SUBAPPLICATION logiBUS_PI_Speed_Publish_OPC (* logiBUS_PI_IDA (Puls-Eingang) als Frequenz (Hz, nur lokal fuer Dashboard/Diagnose) UND als bereits auf die physikalische Einheit umgerechneter Endwert (SCALE+RASTER, M2M-Publish fuer andere Stationen) ausgeben - OHNE jegliche VT-Interaktion. Erweiterung von logiBUS_PI_Raw_Publish_OPC um die Hz->Einheit-Umrechnung (bisher zentral auf STG1 via AR_HZ_TO_Q_Publish_OPC) - jetzt co-located mit dem Sensor: nur der fertige physikalische Endwert verlaesst die Station M2M, der rohe Hz-Wert bleibt lokal. *)
  (* Standard: 61499-2; Description: Copyright (c) 2026 Meisterschulen am Ostbahnhof This program and the accompanying materials are made available under the terms of the Eclipse Public License 2.0 which is available at https://www.eclipse.org/legal/epl-2.0/ SPDX-License-Identifier: EPL-2.0 *)
  (* Version 1.3, 2026-10-03, Franz Höpfinger, Meisterschulen am Ostbahnhof, Franz: 'K auch auf Adapter umstellen' - FT_DERIV_10_AR.K ist jetzt selbst ein AUI-Adapter-Socket (FT_DERIV_10_AR v1.2), die bisherige Entpack-Umgehung ToUINT (AUI_UI_TO_UINT) entfaellt dadurch ersatzlos: ToAUI.AUI_OUT verdrahtet jetzt direkt auf FT_DERIV_10_AR.K (beides AUI-Adapter). *)
  (* Version 1.2, 2026-10-03, Franz Höpfinger, Meisterschulen am Ostbahnhof, Franz: FT_DERIV_10_AR.K (Fensterbreite 0-9, bisher Parameter=9 fest) soll per INI/Dashboard einstellbar sein, 'wie es FilterTimeS auch schon ist'. Neue DerivK/INI_DerivK (gleiches Muster wie FilterTimeS/INI_FilterTimeS, gleiche sSection, eigener KEY='DerivK', Default REAL#9.0) + ToAUI/ToUINT (AR_TO_AUI + neues AUI_UI_TO_UINT, entpackt den Adapter-Wert in eine echte plain UINT-Variable fuer FT_DERIV_10_AR.K - direktes .D1-Dot-Access eines fremden Plugs in eine nicht-adapter-native InputVar wuerde einen 4diac-IDE-Typfehler verursachen, den validate_sub.py nicht sieht, siehe iec61499-creator-Skill). stObjDerivK bleibt wie stObjFilterTimeS auf ID_NULL (kein VT-Eingabefeld platziert, reine Dashboard/INI-Einstellung). Gilt automatisch fuer alle 5 Sensoren, die diesen gemeinsamen Baustein nutzen. *)
  (* Version 1.1, 2026-10-03, Franz Höpfinger, Meisterschulen am Ostbahnhof, Auf Funktionsstand von logiBUS_PI_Raw_Publish_OPC v1.2 gehoben (war seit v1.0 nicht mitgezogen worden) + SCALE/RASTER-Migration fuer alle 5 Puls-Sensoren (Aufnahme B03, Igelband1/2 B10/B11, Zapfwelle B21, Saegeblatt B08): FilterTimeS/INI_FilterTimeS/AR_S_TO_ATM (einstellbare+INI-persistierte PT1-Filterzeit, siehe v1.1 dort) uebernommen, hartcodierten initval_ATM(T#2s) entfernt. Neuer RASTER-InputVar + ROUND_STEP_AR (Round_Final) rundet den FERTIGEN physikalischen Wert NACH der SCALE-Multiplikation (nicht mehr in Hz wie bei logiBUS_PI_Raw_Publish_OPC.RASTER_HZ) - intuitive Werte direkt in der Anzeigeeinheit (z.B. 0.125 U/min, 0.1 km/h) statt der schwer lesbaren Hz-Domaene-Umrechnung. Der lokale Hz-Wert (ID_HZ_WRITE) bleibt bewusst ungerundet, reine Diagnose/Dashboard-Ausgabe, keine andere Station soll ihn remote abonnieren (siehe OPC_UA_NAMENSKONVENTION_LOC_WEB_M2M.md, Scope LOC). *)
  (* Version 1.0, 2026-09-17, Franz Höpfinger, Meisterschulen am Ostbahnhof, initial implementation - Franz: 'die Impulseingaenge will ich auch die Umrechnung auf dem Quellgeraet haben'. Erweitert logiBUS_PI_Raw_Publish_OPC (Rohwert-Kette: logiBUS_PI_IDA -> AD_TO_AR_NUM -> FT_DERIV_10_AR -> FT_PT1_AR, unveraendert) um AR_SPLIT_2 + initval_AR(SCALE) + AR_MUL_2 + zweite AR_PUBLISH_1-Instanz fuer den umgerechneten physikalischen Endwert - analog zum bisherigen AR_HZ_TO_Q_Publish_OPC-Muster (STG1), jetzt aber co-located mit dem Sensor statt zentral. *)
  PACKAGE MyLib::sys;
  IMPORT logiBUS::io::PI::logiBUS_PI;
  IMPORT logiBUS::io::PI::logiBUS_PI_S;
  IMPORT isobus::UT::Q::const::IDs::ID_NULL;
  IMPORT logiBUS::utils::conversion::phys::NumericObjectPool_S;
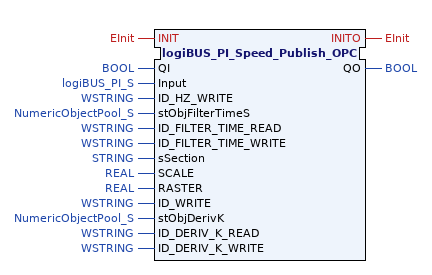
  EVENT_INPUT
    INIT : EInit; (* Initialization Request *)
  END_EVENT
  EVENT_OUTPUT
    INITO : EInit; (* Initialization Confirm *)
  END_EVENT
  VAR_INPUT
    QI : BOOL := TRUE; (* Quality Input - TRUE to enable service *)
    Input : logiBUS::io::PI::logiBUS_PI_S := logiBUS_PI::Invalid; (* Identify the Input PulseInput_I1..I9 *)
    ID_HZ_WRITE : WSTRING; (* Frequenz-Publish-Adresse (REAL Hz, ACTION=PUBLISH), lokal auf dieser Station - nur Dashboard/Diagnose, keine andere Station soll dies remote abonnieren (LOC-Scope) *)
    stObjFilterTimeS : logiBUS::utils::conversion::phys::NumericObjectPool_S := (u16ObjId := ID_NULL, r32Scale := 1.0, i32Offset := 0, u8Decimals := 1); (* Object ID + Scale/Offset/Decimals CNumberVariable (PT1-Filterzeit in Sekunden, VT-Eingabefeld) *)
    ID_FILTER_TIME_READ : WSTRING; (* Remote-Subscribe-Adresse (REAL Sekunden, ACTION=SUBSCRIBE) fuer Web-Override der Filterzeit *)
    ID_FILTER_TIME_WRITE : WSTRING; (* Lokale Echo/Re-Publish-Adresse (REAL Sekunden, ACTION=PUBLISH) der aktuellen Filterzeit *)
    sSection : STRING; (* INI settings.ini Section fuer die persistierte Filterzeit (eindeutig pro Sensor-Instanz) *)
    SCALE : REAL; (* Skalierungsfaktor Hz -> physikalische Einheit (z.B. 3.6/53 fuer km/h, 60.0 fuer U/min bei 1 Impuls/Umdrehung) *)
    RASTER : REAL := 0.001; (* Rundungsraster des FERTIGEN physikalischen Werts (nach SCALE), in der Anzeigeeinheit (z.B. 0.125 fuer U/min, 0.1 fuer km/h) - Platzhalter-Default 0.001 (praktisch kein Runden) *)
    ID_WRITE : WSTRING; (* Publish-Adresse des umgerechneten physikalischen Endwerts (REAL, ACTION=PUBLISH) - das ist die Adresse, die andere Stationen remote abonnieren (M2M-Scope) *)
    stObjDerivK : logiBUS::utils::conversion::phys::NumericObjectPool_S := (u16ObjId := ID_NULL, r32Scale := 1.0, i32Offset := 0, u8Decimals := 0); (* Object ID + Scale/Offset/Decimals CNumberVariable (FT_DERIV_10_AR.K Fensterbreite 0-9, VT-Eingabefeld, 0 Dezimalstellen) - bleibt auf ID_NULL, solange kein VT-Feld platziert ist (reine Dashboard/INI-Einstellung) *)
    ID_DERIV_K_READ : WSTRING; (* Remote-Subscribe-Adresse (REAL, ACTION=SUBSCRIBE) fuer Web-Override von FT_DERIV_10_AR.K *)
    ID_DERIV_K_WRITE : WSTRING; (* Lokale Echo/Re-Publish-Adresse (REAL, ACTION=PUBLISH) des aktuellen FT_DERIV_10_AR.K *)
  END_VAR
  VAR_OUTPUT
    QO : BOOL; (* Quality Output - TRUE if service executed successfully *)
  END_VAR
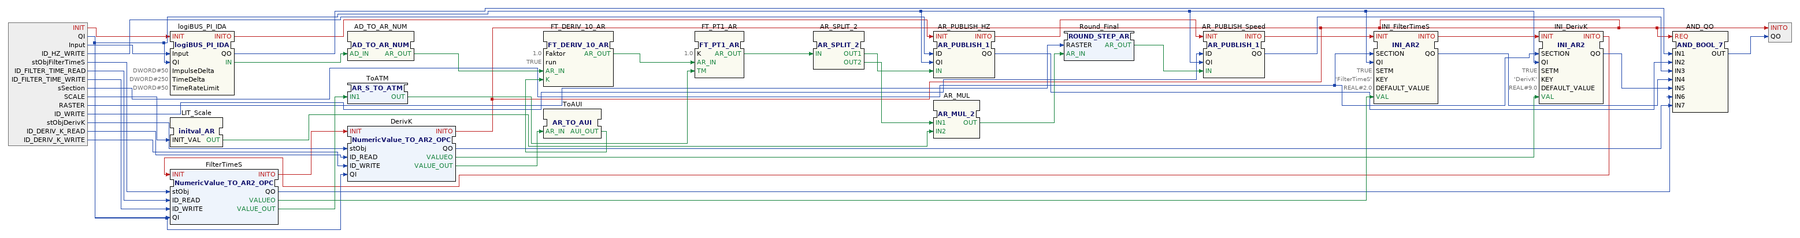
  FBS
    logiBUS_PI_IDA : logiBUS::io::PI::logiBUS_PI_IDA(ImpulseDelta := DWORD#50, TimeDelta := DWORD#250, TimeRateLimit := DWORD#50);
    AD_TO_AR_NUM : adapter::conversion::unidirectional::AD_TO_AR_NUM;
    FT_DERIV_10_AR : OSCAT_adapter::Control::FT_DERIV_10_AR(Faktor := 1.0, run := TRUE);
    FT_PT1_AR : OSCAT_adapter::Control::FT_PT1_AR(K := 1.0);
    AR_SPLIT_2 : adapter::events::unidirectional::AR_SPLIT_2;
    AR_PUBLISH_HZ : adapter::net::AR_PUBLISH_1;
    LIT_Scale : adapter::types::unidirectional::AR::initval::initval_AR;
    AR_MUL : adapter::iec61131::arithmetic::AR_MUL_2;
    AR_PUBLISH_Speed : adapter::net::AR_PUBLISH_1;
    INI_FilterTimeS : eclipse4diac::storage::INI_AR2(SETM := TRUE, KEY := 'FilterTimeS', DEFAULT_VALUE := REAL#2.0);
    INI_DerivK : eclipse4diac::storage::INI_AR2(SETM := TRUE, KEY := 'DerivK', DEFAULT_VALUE := REAL#9.0);
    ToAUI : adapter::conversion::unidirectional::AR_TO_AUI;
    AND_QO : iec61131::booleanOperators::AND_BOOL_7;
  END_FBS
  SUBAPPS
    Round_Final : OSCAT_adapter::Mathematical::ROUND_STEP_AR;
    FilterTimeS : MyLib::sys::NumericValue_TO_AR2_OPC;
    ToATM : MyLib::sys::AR_S_TO_ATM;
    DerivK : MyLib::sys::NumericValue_TO_AR2_OPC;
  END_SUBAPPS
  EVENT_CONNECTIONS
    INIT TO logiBUS_PI_IDA.INIT;
    logiBUS_PI_IDA.INITO TO AR_PUBLISH_HZ.INIT;
    AR_PUBLISH_HZ.INITO TO AR_PUBLISH_Speed.INIT;
    AR_PUBLISH_Speed.INITO TO INI_FilterTimeS.INIT;
    INI_FilterTimeS.INITO TO INI_DerivK.INIT;
    INI_DerivK.INITO TO FilterTimeS.INIT;
    FilterTimeS.INITO TO DerivK.INIT;
    DerivK.INITO TO INITO;
    DerivK.INITO TO AND_QO.REQ;
  END_CONNECTIONS
  DATA_CONNECTIONS
    Input TO logiBUS_PI_IDA.Input;
    ID_HZ_WRITE TO AR_PUBLISH_HZ.ID;
    stObjFilterTimeS TO FilterTimeS.stObj;
    ID_FILTER_TIME_READ TO FilterTimeS.ID_READ;
    ID_FILTER_TIME_WRITE TO FilterTimeS.ID_WRITE;
    sSection TO INI_FilterTimeS.SECTION;
    SCALE TO LIT_Scale.INIT_VAL;
    RASTER TO Round_Final.RASTER;
    ID_WRITE TO AR_PUBLISH_Speed.ID;
    stObjDerivK TO DerivK.stObj;
    ID_DERIV_K_READ TO DerivK.ID_READ;
    ID_DERIV_K_WRITE TO DerivK.ID_WRITE;
    sSection TO INI_DerivK.SECTION;
    QI TO logiBUS_PI_IDA.QI;
    QI TO AR_PUBLISH_HZ.QI;
    QI TO AR_PUBLISH_Speed.QI;
    QI TO INI_FilterTimeS.QI;
    QI TO INI_DerivK.QI;
    logiBUS_PI_IDA.QO TO AND_QO.IN1;
    AR_PUBLISH_HZ.QO TO AND_QO.IN2;
    AR_PUBLISH_Speed.QO TO AND_QO.IN3;
    INI_FilterTimeS.QO TO AND_QO.IN4;
    INI_DerivK.QO TO AND_QO.IN5;
    AND_QO.OUT TO QO;
    QI TO FilterTimeS.QI;
    QI TO DerivK.QI;
    FilterTimeS.QO TO AND_QO.IN6;
    DerivK.QO TO AND_QO.IN7;
  END_CONNECTIONS
  ADAPTER_CONNECTIONS
    logiBUS_PI_IDA.IN TO AD_TO_AR_NUM.AD_IN;
    AD_TO_AR_NUM.AR_OUT TO FT_DERIV_10_AR.AR_IN;
    FT_DERIV_10_AR.AR_OUT TO FT_PT1_AR.AR_IN;
    FilterTimeS.VALUEO TO INI_FilterTimeS.VAL;
    FilterTimeS.VALUE_OUT TO ToATM.IN1;
    ToATM.OUT TO FT_PT1_AR.TM;
    FT_PT1_AR.AR_OUT TO AR_SPLIT_2.IN;
    AR_SPLIT_2.OUT1 TO AR_PUBLISH_HZ.IN;
    AR_SPLIT_2.OUT2 TO AR_MUL.IN1;
    LIT_Scale.OUT TO AR_MUL.IN2;
    AR_MUL.OUT TO Round_Final.AR_IN;
    Round_Final.AR_OUT TO AR_PUBLISH_Speed.IN;
    DerivK.VALUEO TO INI_DerivK.VAL;
    DerivK.VALUE_OUT TO ToAUI.AR_IN;
    ToAUI.AUI_OUT TO FT_DERIV_10_AR.K;
  END_CONNECTIONS
END_SUBAPPLICATION
